(* IEC 61131-3 sources: sis-interlock-demo/src/POUs/PRG_Main, 2 files *)

(* ---- PRG_Main.decl.st ---- *)
// Назначение: главная программа (MainTask, 20 мс): вызывает программу ПАЗ PRG_Sis, которую cemgen
//             генерирует по матрице причин и следствий. В демо без ввода-вывода
//             (GVL_Const.DEMO_IO_SIMULATION) в первом цикле ставит нормальные значения входов:
//             после старта ПЛК все следствия сработали и ждут сброса оператором (раздел 6.10).
// Автор:      kr0nsch
// Версия:     0.1.0
// Документ:   docs/DESIGN.md, раздел «8.4 PRG_Main»
// ВНИМАНИЕ:   код демонстрационный и не предназначен для систем безопасности. Реальная ПАЗ
//             требует определения SIL, сертифицированных аппаратных и программных средств
//             и валидации по ГОСТ Р МЭК 61511.
PROGRAM PRG_Main
VAR
    xFirstCycle : BOOL := TRUE;             // первый цикл после загрузки или старта ПЛК
END_VAR

(* ---- PRG_Main.impl.st ---- *)
// в демо без ввода-вывода — нормальные значения входов в первом цикле
IF xFirstCycle AND GVL_Const.DEMO_IO_SIMULATION THEN
    F_SisIoNormal(stIo := GVL_SisIo.stIo);
END_IF
xFirstCycle := FALSE;
PRG_Sis();
